(* CODESYS project visu_v2.export

Project tree, tasks and I/O mapping:
  visualisation Visu_IOL_O5D150
*)

// /Visu_IOL_O5D150
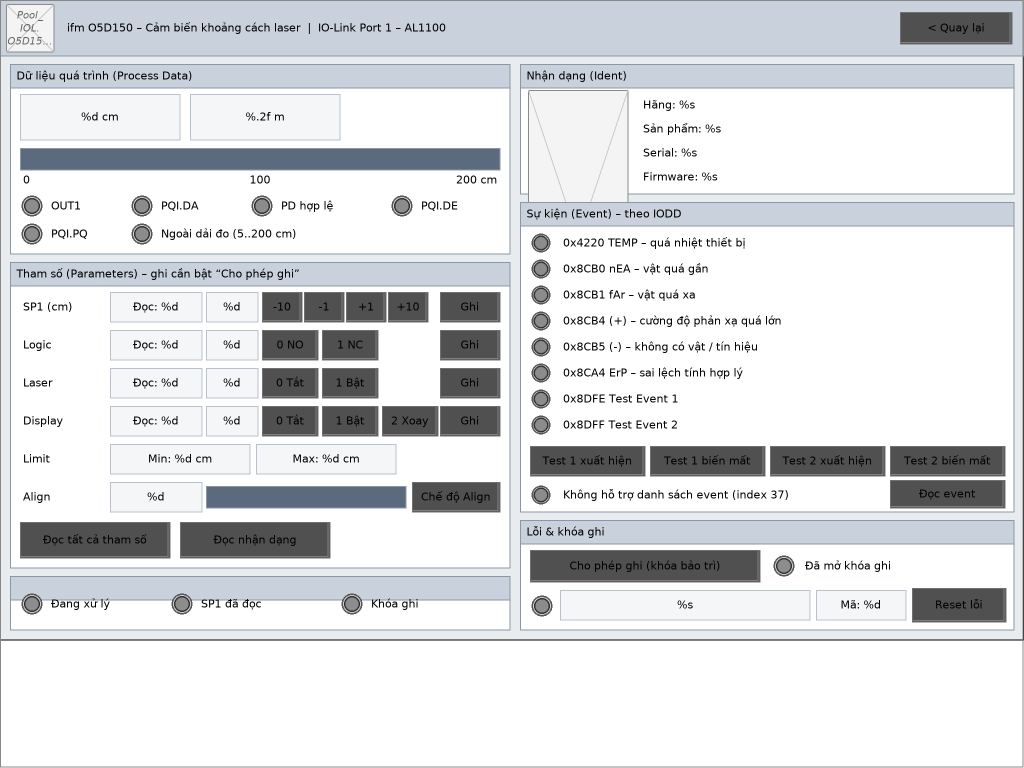
VISUALIZATION Visu_IOL_O5D150  // 1024x768
    Rectangle (0,0 1024x640)
    Rectangle (0,0 1024x56)
    Image (6,4 48x48), image: Pool_IOL.O5D150_icon
    Rectangle (64,0 760x56), "ifm O5D150 – Cảm biến khoảng cách laser | IO-Link Port 1 – AL1100"
    Button (900,12 112x32), "< Quay lại"
        OnMouseClick:  Assign=Visu_Main, Type=Assignment
    Rectangle (10,64 500x190)
    Rectangle (10,64 500x24), "Dữ liệu quá trình (Process Data)"
    Rectangle (20,94 160x46), "%d cm", text variable: GVL_HMI_IOL.stO5D150.uiDistance_cm
    Rectangle (190,94 150x46), "%.2f m", text variable: GVL_HMI_IOL.stO5D150.rDistance_m
    Rectangle (20,148 480x22)
    Rectangle (20,148 480x22)
        p874137650: -(480 - MIN(480, UINT_TO_INT(GVL_HMI_IOL.stO5D150.uiDistance_cm) * 480 / 200))
    Rectangle (20,172 60x16), "0"
    Rectangle (230,172 60x16), "100"
    Rectangle (440,172 60x16), "200 cm"
    Lamp1 (20,194 24x24), variable: GVL_HMI_IOL.stO5D150.xOut1, style: Lamp-Lamp1-Gray
    Rectangle (48,194 60x24), "OUT1"
    Lamp1 (130,194 24x24), variable: GVL_HMI_IOL.stO5D150.xDA, style: Lamp-Lamp1-Gray
    Rectangle (158,194 70x24), "PQI.DA"
    Lamp1 (250,194 24x24), variable: GVL_HMI_IOL.stO5D150.xPdValid, style: Lamp-Lamp1-Gray
    Rectangle (278,194 90x24), "PD hợp lệ"
    Lamp1 (390,194 24x24), variable: GVL_HMI_IOL.stO5D150.xDE, style: Lamp-Lamp1-Gray
    Rectangle (418,194 80x24), "PQI.DE"
    Lamp1 (20,222 24x24), variable: GVL_HMI_IOL.stO5D150.xPQ, style: Lamp-Lamp1-Gray
    Rectangle (48,222 70x24), "PQI.PQ"
    Lamp1 (130,222 24x24), variable: GVL_HMI_IOL.stO5D150.xOutOfRange, style: Lamp-Lamp1-Gray
    Rectangle (158,222 220x24), "Ngoài dải đo (5..200 cm)"
    Rectangle (10,262 500x306)
    Rectangle (10,262 500x24), "Tham số (Parameters) – ghi cần bật “Cho phép ghi”"
    Rectangle (20,292 90x30), "SP1 (cm)"
    Rectangle (110,292 92x30), "Đọc: %d", text variable: GVL_HMI_IOL.stO5D150.uiSP1
    Rectangle (206,292 52x30), "%d", text variable: GVL_HMI_IOL.stO5D150.uiSetSP1
    Button (262,292 40x30), "-10", input disabled if: NOT GVL_HMI_IOL.xMaintEnable
        OnMouseClick: execute { GVL_HMI_IOL.stO5D150.uiSetSP1 := DINT_TO_UINT(LIMIT(5, UINT_TO_DINT(GVL_HMI_IOL.stO5D150.uiSetSP1) + (-10), 200)); }
    Button (304,292 40x30), "-1", input disabled if: NOT GVL_HMI_IOL.xMaintEnable
        OnMouseClick: execute { GVL_HMI_IOL.stO5D150.uiSetSP1 := DINT_TO_UINT(LIMIT(5, UINT_TO_DINT(GVL_HMI_IOL.stO5D150.uiSetSP1) + (-1), 200)); }
    Button (346,292 40x30), "+1", input disabled if: NOT GVL_HMI_IOL.xMaintEnable
        OnMouseClick: execute { GVL_HMI_IOL.stO5D150.uiSetSP1 := DINT_TO_UINT(LIMIT(5, UINT_TO_DINT(GVL_HMI_IOL.stO5D150.uiSetSP1) + (1), 200)); }
    Button (388,292 40x30), "+10", input disabled if: NOT GVL_HMI_IOL.xMaintEnable
        OnMouseClick: execute { GVL_HMI_IOL.stO5D150.uiSetSP1 := DINT_TO_UINT(LIMIT(5, UINT_TO_DINT(GVL_HMI_IOL.stO5D150.uiSetSP1) + (10), 200)); }
    Button (440,292 60x30), "Ghi", input disabled if: NOT GVL_HMI_IOL.xMaintEnable
        OnMouseClick: execute { GVL_HMI_IOL.stO5D150.xCmdWriteSP1 := TRUE; }
    Rectangle (20,330 90x30), "Logic"
    Rectangle (110,330 92x30), "Đọc: %d", text variable: GVL_HMI_IOL.stO5D150.usiLogic
    Rectangle (206,330 52x30), "%d", text variable: GVL_HMI_IOL.stO5D150.usiSetLogic
    Button (262,330 56x30), "0 NO", input disabled if: NOT GVL_HMI_IOL.xMaintEnable
        OnMouseClick: execute { GVL_HMI_IOL.stO5D150.usiSetLogic := 0; }
    Button (322,330 56x30), "1 NC", input disabled if: NOT GVL_HMI_IOL.xMaintEnable
        OnMouseClick: execute { GVL_HMI_IOL.stO5D150.usiSetLogic := 1; }
    Button (440,330 60x30), "Ghi", input disabled if: NOT GVL_HMI_IOL.xMaintEnable
        OnMouseClick: execute { GVL_HMI_IOL.stO5D150.xCmdWriteLogic := TRUE; }
    Rectangle (20,368 90x30), "Laser"
    Rectangle (110,368 92x30), "Đọc: %d", text variable: GVL_HMI_IOL.stO5D150.usiLaser
    Rectangle (206,368 52x30), "%d", text variable: GVL_HMI_IOL.stO5D150.usiSetLaser
    Button (262,368 56x30), "0 Tắt", input disabled if: NOT GVL_HMI_IOL.xMaintEnable
        OnMouseClick: execute { GVL_HMI_IOL.stO5D150.usiSetLaser := 0; }
    Button (322,368 56x30), "1 Bật", input disabled if: NOT GVL_HMI_IOL.xMaintEnable
        OnMouseClick: execute { GVL_HMI_IOL.stO5D150.usiSetLaser := 1; }
    Button (440,368 60x30), "Ghi", input disabled if: NOT GVL_HMI_IOL.xMaintEnable
        OnMouseClick: execute { GVL_HMI_IOL.stO5D150.xCmdWriteLaser := TRUE; }
    Rectangle (20,406 90x30), "Display"
    Rectangle (110,406 92x30), "Đọc: %d", text variable: GVL_HMI_IOL.stO5D150.usiDisplay
    Rectangle (206,406 52x30), "%d", text variable: GVL_HMI_IOL.stO5D150.usiSetDisplay
    Button (262,406 56x30), "0 Tắt", input disabled if: NOT GVL_HMI_IOL.xMaintEnable
        OnMouseClick: execute { GVL_HMI_IOL.stO5D150.usiSetDisplay := 0; }
    Button (322,406 56x30), "1 Bật", input disabled if: NOT GVL_HMI_IOL.xMaintEnable
        OnMouseClick: execute { GVL_HMI_IOL.stO5D150.usiSetDisplay := 1; }
    Button (382,406 56x30), "2 Xoay", input disabled if: NOT GVL_HMI_IOL.xMaintEnable
        OnMouseClick: execute { GVL_HMI_IOL.stO5D150.usiSetDisplay := 2; }
    Button (440,406 60x30), "Ghi", input disabled if: NOT GVL_HMI_IOL.xMaintEnable
        OnMouseClick: execute { GVL_HMI_IOL.stO5D150.xCmdWriteDisplay := TRUE; }
    Rectangle (20,444 90x30), "Limit"
    Rectangle (110,444 140x30), "Min: %d cm", text variable: GVL_HMI_IOL.stO5D150.uiLimitMin_cm
    Rectangle (256,444 140x30), "Max: %d cm", text variable: GVL_HMI_IOL.stO5D150.uiLimitMax_cm
    Rectangle (20,482 90x30), "Align"
    Rectangle (110,482 92x30), "%d", text variable: GVL_HMI_IOL.stO5D150.usiAlign
    Rectangle (206,486 200x22)
    Rectangle (206,486 200x22)
        p874137650: -(200 - MIN(200, USINT_TO_INT(GVL_HMI_IOL.stO5D150.usiAlign) * 200 / 100))
    Button (412,482 88x30), "Chế độ Align"
        OnMouseClick: execute { GVL_HMI_IOL.stO5D150.xAlignMode := NOT GVL_HMI_IOL.stO5D150.xAlignMode; }
    Button (20,522 150x36), "Đọc tất cả tham số"
        OnMouseClick: execute { GVL_HMI_IOL.stO5D150.xCmdReadAll := TRUE; }
    Button (180,522 150x36), "Đọc nhận dạng"
        OnMouseClick: execute { GVL_HMI_IOL.stO5D150.xCmdReadIdent := TRUE; }
    Rectangle (10,576 500x54)
    Rectangle (10,576 500x24)
    Lamp1 (20,592 24x24), variable: GVL_HMI_IOL.stO5D150.xBusy, style: Lamp-Lamp1-Gray
    Rectangle (48,592 110x24), "Đang xử lý"
    Lamp1 (170,592 24x24), variable: GVL_HMI_IOL.stO5D150.xParamValid, style: Lamp-Lamp1-Gray
    Rectangle (198,592 130x24), "SP1 đã đọc"
    Lamp1 (340,592 24x24), variable: GVL_HMI_IOL.stO5D150.xWriteLocked, style: Lamp-Lamp1-Gray
    Rectangle (368,592 130x24), "Khóa ghi"
    Rectangle (520,64 494x130)
    Rectangle (520,64 494x24), "Nhận dạng (Ident)"
    Image (528,90 100x300), image: Pool_IOL.O5D150_pic
    Rectangle (640,94 366x22), "Hãng: %s", text variable: GVL_HMI_IOL.stO5D150.sVendor
    Rectangle (640,118 366x22), "Sản phẩm: %s", text variable: GVL_HMI_IOL.stO5D150.sProduct
    Rectangle (640,142 366x22), "Serial: %s", text variable: GVL_HMI_IOL.stO5D150.sSerial
    Rectangle (640,166 366x22), "Firmware: %s", text variable: GVL_HMI_IOL.stO5D150.sFwRev
    Rectangle (520,202 494x310)
    Rectangle (520,202 494x24), "Sự kiện (Event) – theo IODD"
    Lamp1 (530,232 22x22), variable: GVL_HMI_IOL.stO5D150.axEvtActive[0], style: Lamp-Lamp1-Gray
    Rectangle (560,231 440x24), "0x4220 TEMP – quá nhiệt thiết bị"
    Lamp1 (530,258 22x22), variable: GVL_HMI_IOL.stO5D150.axEvtActive[1], style: Lamp-Lamp1-Gray
    Rectangle (560,257 440x24), "0x8CB0 nEA – vật quá gần"
    Lamp1 (530,284 22x22), variable: GVL_HMI_IOL.stO5D150.axEvtActive[2], style: Lamp-Lamp1-Gray
    Rectangle (560,283 440x24), "0x8CB1 fAr – vật quá xa"
    Lamp1 (530,310 22x22), variable: GVL_HMI_IOL.stO5D150.axEvtActive[3], style: Lamp-Lamp1-Gray
    Rectangle (560,309 440x24), "0x8CB4 (+) – cường độ phản xạ quá lớn"
    Lamp1 (530,336 22x22), variable: GVL_HMI_IOL.stO5D150.axEvtActive[4], style: Lamp-Lamp1-Gray
    Rectangle (560,335 440x24), "0x8CB5 (-) – không có vật / tín hiệu"
    Lamp1 (530,362 22x22), variable: GVL_HMI_IOL.stO5D150.axEvtActive[5], style: Lamp-Lamp1-Gray
    Rectangle (560,361 440x24), "0x8CA4 ErP – sai lệch tính hợp lý"
    Lamp1 (530,388 22x22), variable: GVL_HMI_IOL.stO5D150.axEvtActive[6], style: Lamp-Lamp1-Gray
    Rectangle (560,387 440x24), "0x8DFE Test Event 1"
    Lamp1 (530,414 22x22), variable: GVL_HMI_IOL.stO5D150.axEvtActive[7], style: Lamp-Lamp1-Gray
    Rectangle (560,413 440x24), "0x8DFF Test Event 2"
    Button (530,446 115x30), "Test 1 xuất hiện", input disabled if: NOT GVL_HMI_IOL.xMaintEnable
        OnMouseClick: execute { GVL_HMI_IOL.stO5D150.xCmdTestEvt1On := TRUE; }
    Button (650,446 115x30), "Test 1 biến mất", input disabled if: NOT GVL_HMI_IOL.xMaintEnable
        OnMouseClick: execute { GVL_HMI_IOL.stO5D150.xCmdTestEvt1Off := TRUE; }
    Button (770,446 115x30), "Test 2 xuất hiện", input disabled if: NOT GVL_HMI_IOL.xMaintEnable
        OnMouseClick: execute { GVL_HMI_IOL.stO5D150.xCmdTestEvt2On := TRUE; }
    Button (890,446 115x30), "Test 2 biến mất", input disabled if: NOT GVL_HMI_IOL.xMaintEnable
        OnMouseClick: execute { GVL_HMI_IOL.stO5D150.xCmdTestEvt2Off := TRUE; }
    Lamp1 (530,484 22x22), variable: GVL_HMI_IOL.stO5D150.xEvtListNotSupported, style: Lamp-Lamp1-Gray
    Rectangle (560,483 320x24), "Không hỗ trợ danh sách event (index 37)"
    Button (890,480 115x28), "Đọc event"
        OnMouseClick: execute { GVL_HMI_IOL.stO5D150.xCmdReadEvents := TRUE; }
    Rectangle (520,520 494x110)
    Rectangle (520,520 494x24), "Lỗi & khóa ghi"
    Button (530,550 230x32), "Cho phép ghi (khóa bảo trì)"
        OnMouseClick: execute { GVL_HMI_IOL.xMaintEnable := NOT GVL_HMI_IOL.xMaintEnable; }
    Lamp1 (772,554 24x24), variable: GVL_HMI_IOL.xMaintEnable, style: Lamp-Lamp1-Gray
    Rectangle (802,554 200x24), "Đã mở khóa ghi"
    Lamp1 (530,594 24x24), variable: GVL_HMI_IOL.stO5D150.xError, style: Lamp-Lamp1-Gray
    Rectangle (560,590 250x30), "%s", text variable: GVL_HMI_IOL.stO5D150.wsErrText
    Rectangle (816,590 90x30), "Mã: %d", text variable: GVL_HMI_IOL.stO5D150.uiDevErr
    Button (912,588 94x34), "Reset lỗi"
        OnMouseClick: execute { GVL_HMI_IOL.stO5D150.xCmdResetErr := TRUE; }
END_VISUALIZATION
